(* IEC 61131-3 sources: llm-plc-st-eval/data/definitivo/qwen2.5-coder_14b/I8/zero_shot, 3 files *)

(* ---- ejec_1.st ---- *)
```pascal
FUNCTION_BLOCK FB_Compresor
VAR_INPUT
    pOilOk : BOOL; // Presión de aceite correcta
    tempOk : BOOL; // Temperatura correcta
    sinAlm : BOOL; // Ausencia de alarmas
    btnMarcha : BOOL; // Botón de marcha
    btnParo : BOOL; // Botón de paro
END_VAR

VAR_OUTPUT
    comp : BOOL; // Salida del compresor
    causaBloqueo : INT; // Causa del bloqueo
END_VAR

VAR
    timerOilOk : TON; // Temporizador para la presión de aceite
    marchaAnterior : BOOL; // Estado anterior del botón de marcha
    paroAnterior : BOOL; // Estado anterior del botón de paro
    permisivoCumplido : BOOL; // Indica si todos los permisivos están cumplidos
    estadoMarcha : BOOL; // Estado actual del compresor
END_VAR

// Inicialización del temporizador
IF NOT timerOilOk.Q THEN
    timerOilOk(IN := FALSE, PT := T#3S);
END_IF;

// Actualización de estados anteriores
marchaAnterior := btnMarcha;
paroAnterior := btnParo;

// Lógica de paro
IF btnParo AND NOT paroAnterior THEN
    comp := FALSE;
    estadoMarcha := FALSE;
END_IF;

// Lógica de arranque
IF btnMarcha AND NOT marchaAnterior THEN
    timerOilOk(IN := pOilOk);
    permisivoCumplido := pOilOk AND tempOk AND sinAlm;
    IF permisivoCumplido THEN
        comp := TRUE;
        estadoMarcha := TRUE;
    END_IF;
END_IF;

// Mantener el compresor en marcha si ya está arrancado
IF estadoMarcha THEN
    comp := TRUE;
ELSE
    comp := FALSE;
END_IF;

// Determinar la causa del bloqueo
IF NOT pOilOk THEN
    causaBloqueo := 1;
ELSIF NOT tempOk THEN
    causaBloqueo := 2;
ELSIF NOT sinAlm THEN
    causaBloqueo := 3;
ELSE
    causaBloqueo := 0;
END_IF;

// Reiniciar el temporizador si la presión de aceite se pierde
IF NOT pOilOk THEN
    timerOilOk(IN := FALSE);
END_IF;

END_FUNCTION_BLOCK
```

(* ---- ejec_2.st ---- *)
```pascal
FUNCTION_BLOCK FB_Compresor
VAR_INPUT
    pOilOk : BOOL; // Presión de aceite correcta
    tempOk : BOOL; // Temperatura correcta
    sinAlm : BOOL; // Ausencia de alarmas
    btnMarcha : BOOL; // Botón de marcha
    btnParo : BOOL; // Botón de paro
END_VAR

VAR_OUTPUT
    comp : BOOL; // Salida del compresor
    causaBloqueo : INT; // Causa de bloqueo
END_VAR

VAR
    timerOilOk : TON; // Temporizador para presión de aceite
    marchaAnterior : BOOL; // Estado anterior del botón de marcha
    paroAnterior : BOOL; // Estado anterior del botón de paro
    permisivoCumplido : BOOL; // Indica si se cumplen todos los permisivos
END_VAR

// Inicialización del temporizador
IF NOT timerOilOk.Q THEN
    timerOilOk(IN := FALSE, PT := T#3S);
END_IF

// Detectar transición de botón de marcha
IF btnMarcha AND NOT marchaAnterior THEN
    timerOilOk(IN := pOilOk);
END_IF

// Detectar transición de botón de paro
IF btnParo AND NOT paroAnterior THEN
    comp := FALSE;
END_IF

// Actualizar estado de botones
marchaAnterior := btnMarcha;
paroAnterior := btnParo;

// Verificar permisivos
permisivoCumplido := pOilOk AND tempOk AND sinAlm AND timerOilOk.Q;

// Determinar causa de bloqueo
IF NOT pOilOk THEN
    causaBloqueo := 1;
ELSIF NOT tempOk THEN
    causaBloqueo := 2;
ELSIF NOT sinAlm THEN
    causaBloqueo := 3;
ELSE
    causaBloqueo := 0;
END_IF

// Control de arranque y paro
IF btnParo THEN
    comp := FALSE;
ELSEIF btnMarcha AND permisivoCumplido THEN
    comp := TRUE;
END_IF
END_FUNCTION_BLOCK
```

(* ---- ejec_3.st ---- *)
```pascal
FUNCTION_BLOCK FB_Compresor
VAR_INPUT
    pOilOk : BOOL; // Presión de aceite correcta
    tempOk : BOOL; // Temperatura correcta
    sinAlm : BOOL; // Ausencia de alarmas
    btnMarcha : BOOL; // Botón de marcha
    btnParo : BOOL; // Botón de paro
END_VAR

VAR_OUTPUT
    comp : BOOL; // Salida del compresor
    causaBloqueo : INT; // Causa de bloqueo
END_VAR

VAR
    timerOilOk : TON; // Temporizador para presión de aceite
    estadoMarcha : BOOL; // Estado de marcha del compresor
    lastBtnMarcha : BOOL; // Estado anterior del botón de marcha
    lastBtnParo : BOOL; // Estado anterior del botón de paro
END_VAR

// Inicialización
IF NOT estadoMarcha THEN
    comp := FALSE;
    causaBloqueo := 0;
END_IF

// Actualización de estados de botones
IF btnMarcha <> lastBtnMarcha THEN
    lastBtnMarcha := btnMarcha;
END_IF

IF btnParo <> lastBtnParo THEN
    lastBtnParo := btnParo;
END_IF

// Paro del compresor por botón de paro o pérdida de permisivos
IF btnParo OR (estadoMarcha AND (NOT pOilOk OR NOT tempOk OR NOT sinAlm)) THEN
    comp := FALSE;
    estadoMarcha := FALSE;
END_IF

// Inicio del compresor por botón de marcha
IF NOT estadoMarcha AND btnMarcha AND pOilOk AND tempOk AND sinAlm THEN
    comp := TRUE;
    estadoMarcha := TRUE;
END_IF

// Control de la causa de bloqueo
IF NOT pOilOk THEN
    causaBloqueo := 1;
ELSIF NOT tempOk THEN
    causaBloqueo := 2;
ELSIF NOT sinAlm THEN
    causaBloqueo := 3;
ELSE
    causaBloqueo := 0;
END_IF

// Temporizador para presión de aceite
timerOilOk(IN := pOilOk, PT := T#3S);
IF timerOilOk.Q THEN
    // Presión de aceite correcta durante 3 segundos
    // (No se necesita acción adicional aquí)
END_IF

END_FUNCTION_BLOCK
```
